PROGRAM PRG_Tests
{IF defined (S85_PROD)}
{IF defined (S85_TEST_BUILD)}
{error 'S85_PROD and S85_TEST_BUILD cannot both be defined'}
{END_IF}
{END_IF}
VAR
{IF defined (S85_TEST_BUILD)}
    fbLightTests : FB_LightTests;
    fbButtonTests : FB_ButtonTests;
    fbLightCatalogTests : FB_LightCatalogTests;
    fbLocationWorkshopTests : FB_Location_WorkshopTests;
    fbMqttLightBuilderTests : FB_MqttLightBuilderTests;
    fbMqttLightProtocolTests : FB_MqttLightProtocolTests;
    fbMqttCanaryParserTests : FB_MqttCanaryParserTests;
{END_IF}
END_VAR

{IF defined (S85_TEST_BUILD)}
TcUnit.RUN();
{END_IF}

END_PROGRAM

(* stored: Version 1.1.0.1
   POU PRG_Tests: Id {879b7b3f-bff0-4ef4-9304-d849213a653e}, SpecialFunc None *)
